SUBAPPLICATION FU_Skalierung (* H300-Rohwerte (UINT-Register) in physikalische Werte umrechnen. RD_n = Reihenfolge des CLIENT_0_8 in FU_Messwerte, SD_n = Reihenfolge des PUBLISH_8. Die festen Schnittstellentypen (UINT rein, REAL/UINT raus) typisieren die ANY-Pins von CLIENT und PUBLISH. *)
  (* Standard: 61499-2; Description: Copyright (c) 2026 Franz Höpfinger This program and the accompanying materials are made available under the terms of the Eclipse Public License 2.0 which is available at https://www.eclipse.org/legal/epl-2.0/ SPDX-License-Identifier: EPL-2.0 *)
  (* Version 1.0, 2026-11-02, Franz Höpfinger, Franz Höpfinger, aus FU_Messwerte herausgeloest *)
  PACKAGE FBs::FU_Demo;
  IMPORT FBs::FU_Demo::FU_Demo_Konstanten::FU_SKALIERUNG_0_01;
  IMPORT FBs::FU_Demo::FU_Demo_Konstanten::FU_SKALIERUNG_0_1;
  IMPORT FBs::FU_Demo::FU_Demo_Konstanten::FU_SKALIERUNG_1;
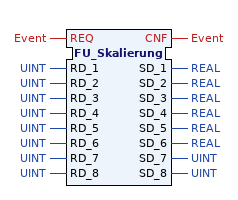
  EVENT_INPUT
    REQ; (* Neue Rohwerte (von CLIENT_0_8.CNF) *)
  END_EVENT
  EVENT_OUTPUT
    CNF; (* Alle Werte umgerechnet *)
  END_EVENT
  VAR_INPUT
    RD_1 : UINT; (* Rohwert 9000H vom Modbus-Client *)
    RD_2 : UINT; (* Rohwert 9001H vom Modbus-Client *)
    RD_3 : UINT; (* Rohwert 9002H vom Modbus-Client *)
    RD_4 : UINT; (* Rohwert 9003H vom Modbus-Client *)
    RD_5 : UINT; (* Rohwert 9004H vom Modbus-Client *)
    RD_6 : UINT; (* Rohwert 9006H vom Modbus-Client *)
    RD_7 : UINT; (* Rohwert 9332H vom Modbus-Client *)
    RD_8 : UINT; (* Rohwert 9333H vom Modbus-Client *)
  END_VAR
  VAR_OUTPUT
    SD_1 : REAL; (* Ist-Frequenz in Hz (9000H) *)
    SD_2 : REAL; (* wirksame Soll-Frequenz in Hz (9001H) *)
    SD_3 : REAL; (* Ausgangsstrom in A (9002H) *)
    SD_4 : REAL; (* Ausgangsspannung in V (9003H) *)
    SD_5 : REAL; (* Zwischenkreisspannung in V (9004H) *)
    SD_6 : REAL; (* Ausgangsleistung in kW (9006H) *)
    SD_7 : UINT; (* Betriebsstatus (9332H): 1=vorwaerts, 2=rueckwaerts, 3=Stopp *)
    SD_8 : UINT; (* Fehlercode (9333H): 0=keine Stoerung *)
  END_VAR
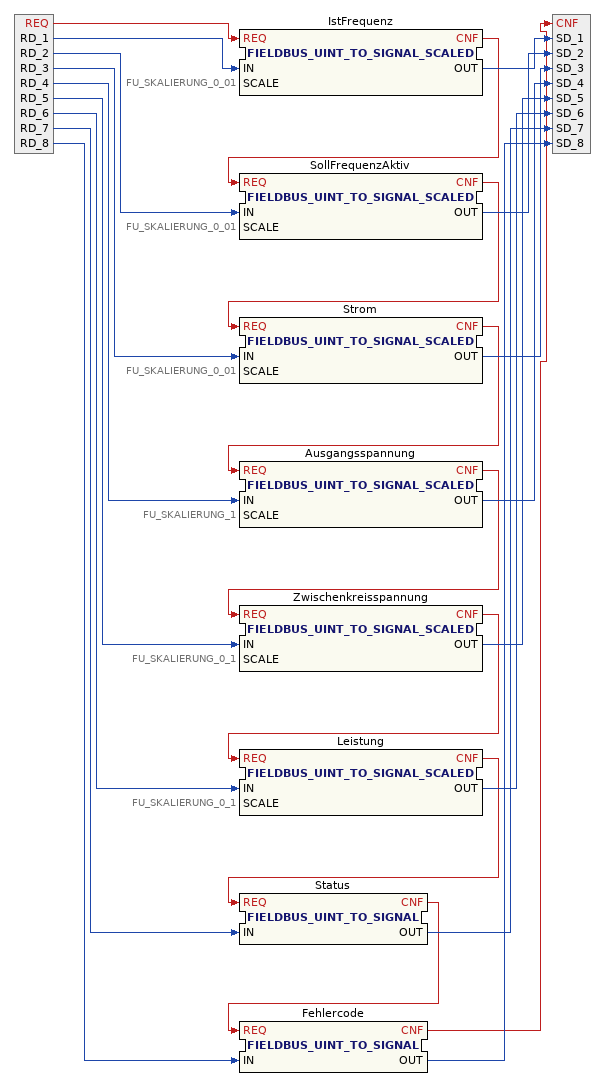
  FBS
    IstFrequenz : logiBUS::signalprocessing::fieldbus::FIELDBUS_UINT_TO_SIGNAL_SCALED(SCALE := FU_SKALIERUNG_0_01); (* 9000H, 0,01 Hz *)
    SollFrequenzAktiv : logiBUS::signalprocessing::fieldbus::FIELDBUS_UINT_TO_SIGNAL_SCALED(SCALE := FU_SKALIERUNG_0_01); (* 9001H, 0,01 Hz - der vom FU tatsaechlich verwendete Sollwert *)
    Strom : logiBUS::signalprocessing::fieldbus::FIELDBUS_UINT_TO_SIGNAL_SCALED(SCALE := FU_SKALIERUNG_0_01); (* 9002H, 0,01 A (Geraete < 75 kW) *)
    Ausgangsspannung : logiBUS::signalprocessing::fieldbus::FIELDBUS_UINT_TO_SIGNAL_SCALED(SCALE := FU_SKALIERUNG_1); (* 9003H, 1 V *)
    Zwischenkreisspannung : logiBUS::signalprocessing::fieldbus::FIELDBUS_UINT_TO_SIGNAL_SCALED(SCALE := FU_SKALIERUNG_0_1); (* 9004H, 0,1 V *)
    Leistung : logiBUS::signalprocessing::fieldbus::FIELDBUS_UINT_TO_SIGNAL_SCALED(SCALE := FU_SKALIERUNG_0_1); (* 9006H, 0,1 kW *)
    Status : logiBUS::signalprocessing::fieldbus::FIELDBUS_UINT_TO_SIGNAL; (* 9332H: 1=Vorwaerts, 2=Rueckwaerts, 3=Stopp *)
    Fehlercode : logiBUS::signalprocessing::fieldbus::FIELDBUS_UINT_TO_SIGNAL; (* 9333H: 0=keine Stoerung, sonst Fehlercode lt. Handbuch 9.1.5.1 *)
  END_FBS
  EVENT_CONNECTIONS
    REQ TO IstFrequenz.REQ;
    IstFrequenz.CNF TO SollFrequenzAktiv.REQ;
    SollFrequenzAktiv.CNF TO Strom.REQ;
    Strom.CNF TO Ausgangsspannung.REQ;
    Ausgangsspannung.CNF TO Zwischenkreisspannung.REQ;
    Zwischenkreisspannung.CNF TO Leistung.REQ;
    Leistung.CNF TO Status.REQ;
    Status.CNF TO Fehlercode.REQ;
    Fehlercode.CNF TO CNF;
  END_CONNECTIONS
  DATA_CONNECTIONS
    RD_1 TO IstFrequenz.IN;
    RD_2 TO SollFrequenzAktiv.IN;
    RD_3 TO Strom.IN;
    RD_4 TO Ausgangsspannung.IN;
    RD_5 TO Zwischenkreisspannung.IN;
    RD_6 TO Leistung.IN;
    RD_7 TO Status.IN;
    RD_8 TO Fehlercode.IN;
    IstFrequenz.OUT TO SD_1;
    SollFrequenzAktiv.OUT TO SD_2;
    Strom.OUT TO SD_3;
    Ausgangsspannung.OUT TO SD_4;
    Zwischenkreisspannung.OUT TO SD_5;
    Leistung.OUT TO SD_6;
    Status.OUT TO SD_7;
    Fehlercode.OUT TO SD_8;
  END_CONNECTIONS
END_SUBAPPLICATION
